{attribute 'qualified_only'}
{attribute 'strict'}
{attribute 'to_string'}
TYPE E_LoggerProviderFailureReason :
(
	NA := 0,  // No failure occurred.
	RECORD_POINTER_NULL,  // The supplied log record pointer is null.
	QUEUE_POP_FAILURE,  // A record could not be popped from the provider's queue during cyclical processing.
	STAGE_PROCESSOR_FAILURE,  // A processor could not be added to the internal linked list for some reason.
	UNEXPECTED_NULL_PROCESSOR_POINTER,  // A processor pointer was invalid when being accessed internally to the provider.
	UNEXPECTED_NULL_LINKED_LIST_NODE  // A processor linked list poitner was invalid when being accessed internally to the provider.
) UDINT;
END_TYPE

(* stored: Version 1.1.0.1
   EnumerationTextList E_LoggerProviderFailureReason: Id {7818a20b-97b0-460d-98a1-374dc1cf8ebe} *)
